{attribute 'Tc2GvlVarNames'}
VAR_GLOBAL
	stgGr01HMI			:ST_Gr01HMIRef;
END_VAR

(* stored: Version 1.1.0.1, ProductVersion 3.1.4024.15
   GVL GVL_Gr01HMI: Id {e1714ec3-ccd1-41b7-b82d-08549a1d2510} *)
